// TIA Portal V21 export
// export: Created 2026-11-11T00:48:11.4062222Z, ExportSetting WithDefaults, DisplayName Totally Integrated Automation Portal, DisplayVersion V21 Update 3, DisplayName STEP 7 Professional, DisplayVersion V21 Update 3, DisplayName STEP 7 Safety, DisplayVersion V21, DisplayName Tech WebApplication, DisplayVersion V21, DisplayName WinCC Basic/Comfort/Advanced, DisplayVersion V21 Update 3, DisplayName WinCC Unified, DisplayVersion V21 Update 3
FUNCTION_BLOCK "FB_Scl_sl019"   // FB48, SCL
{ S7_Optimized_Access := 'TRUE' }
VERSION : 0.1
// stored: AutoNumber true, IsIECCheckEnabled false, IsRetainMemResEnabled false, MemoryReserve 100, SetENOAutomatically false, UDAEnableTagReadback false
   VAR_INPUT
      v_c_no : Counter;
      v_cu : Bool;
      v_cd : Bool;
      v_s : Bool;
      v_pv : Word;
      v_r : Bool;
   END_VAR
   VAR_OUTPUT
      v_q : Bool;
      v_cv : Word;
   END_VAR
BEGIN
   #v_cv := S_CUD(C_NO := #v_c_no, CU := #v_cu, CD := #v_cd, S := #v_s, PV := #v_pv, R := #v_r, Q => #v_q);
END_FUNCTION_BLOCK
